// TIA Portal V20 export
// export: Created 2026-10-19T18:06:56.7145868Z, ExportSetting WithDefaults, DisplayName Totally Integrated Automation Portal, DisplayVersion V20 Update 6, DisplayName TIA Portal Openness, DisplayVersion V20 Update 6, DisplayName TIA Portal Version Control Interface, DisplayVersion V20 Update 6, DisplayName SINAMICS Startdrive Advanced, DisplayVersion V20 SP1, DisplayName SINAMICS Startdrive G130, G150, S120, S150, SINAMICS MV, G220, S200, S210, DisplayVersion V20 SP1, DisplayName SINAMICS Startdrive G110M, G120, G120C, G120D, G120P, G115D, DisplayVersion V20 SP1, DisplayName STEP 7 Professional, DisplayVersion V20 Update 6, DisplayName STEP 7 Safety, DisplayVersion V20 Update 2, DisplayName WinCC Basic/Comfort/Advanced, DisplayVersion V20 Update 6, DisplayName WinCC Unified, DisplayVersion V20 Update 6
DATA_BLOCK "SAI_IND_ZeroAdjust_DB"   // DB111
VERSION : 0.1
// stored: AutoNumber true, DBAccessibleFromOPCUA true, DBAccessibleFromWebserver true, InstanceOfName SAI_IND_ZeroAdjust, InstanceOfType FB
"SAI_IND_ZeroAdjust"
   // VAR_INPUT
   //    ID : HW_IO;
   // END_VAR
   // VAR_OUTPUT
   //    Process : Bool;
   //    Done : Bool;
   //    Error : Bool;
   // END_VAR
   // VAR_IN_OUT
   //    Start : Bool;
   // END_VAR
   // VAR
   //    Activate : Bool;
   //    Status_RECORD : Int;
   //    Zero_RECORD : Int;
   //    WRREC_Zero { S7_SetPoint := 'True'} : WRREC;
   //    RDREC_Status { S7_SetPoint := 'True'} : RDREC;
   //    AdjustStep : SInt;
   //    Static01 : Bool;
   //    Static02 : Bool;
   //    Static03 : Bool;
   // END_VAR
BEGIN
END_DATA_BLOCK
